(* IEC 61131-3 sources: rusty/compiler/plc_cfc/fixtures/blocks/valid/action_bare, 1 file *)

(* ---- counter.st ---- *)
FUNCTION_BLOCK counter
VAR_OUTPUT
    out : DINT;
END_VAR
END_FUNCTION_BLOCK

ACTIONS
    ACTION reset
        out := 0;
    END_ACTION
END_ACTIONS
